SUBAPPLICATION SubApp_PC_A (* Geraet A: Methode AddValues (opcua.adoc): SERVER_1_2 + F_ADD; Input_I1 ruft sie per CLIENT_2_1 mit 43 und 10 auf (Ergebnis 53) *)
  (* Standard: 61499-2; Description: Copyright (c) 2026 Meisterschulen am Ostbahnhof This program and the accompanying materials are made available under the terms of the Eclipse Public License 2.0 which is available at https://www.eclipse.org/legal/epl-2.0/ SPDX-License-Identifier: EPL-2.0 *)
  (* Version 1.0, 2026-10-18, Franz Höpfinger, Meisterschulen am Ostbahnhof, opcua.adoc-Beispiel auf zwei Geraeten *)
  PACKAGE subapp::Training_15_OPC_UA_RES;
  IMPORT VV::const::OPC_UA::myOpcUaAddresses::T15_ADD_CALL;
  IMPORT logiBUS::io::DI::logiBUS_DI::Input_I1;
  IMPORT logiBUS::io::DI::logiBUS_DI_Events::BUTTON_PRESS_DOWN;
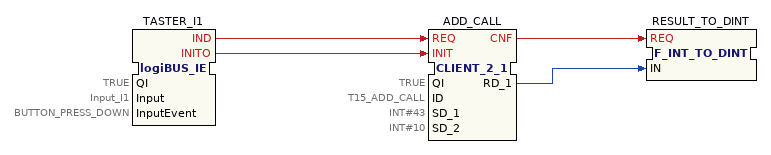
  FBS
    TASTER_I1 : logiBUS::io::DI::logiBUS_IE(QI := TRUE, Input := Input_I1, InputEvent := BUTTON_PRESS_DOWN);
    ADD_CALL : iec61499::net::CLIENT_2_1(QI := TRUE, ID := T15_ADD_CALL, SD_1 := INT#43, SD_2 := INT#10);
    RESULT_TO_DINT : iec61131::conversion::F_INT_TO_DINT;
  END_FBS
  EVENT_CONNECTIONS
    TASTER_I1.IND TO ADD_CALL.REQ;
    TASTER_I1.INITO TO ADD_CALL.INIT;
    ADD_CALL.CNF TO RESULT_TO_DINT.REQ;
  END_CONNECTIONS
  DATA_CONNECTIONS
    ADD_CALL.RD_1 TO RESULT_TO_DINT.IN;
  END_CONNECTIONS
END_SUBAPPLICATION
